// TIA Portal V21 export
TagTable "T_V4"
  X_V4 : Bool  (PLC tag HMI_IF.BtnInit, HMI_Connection_1, 100 ms)
